Fanuc KAREL source: ka00105.KL

-- PROVISIONAL review KL for V940-1; original PC SHA256 45f8fe3be269b6ab01cad793c02046efcd257036997fb4219fc5ec4bbcc30542
-- Incomplete behavior may be omitted. Consult companion uncertainty JSON. Do not deploy.
PROGRAM KA00105
%NOLOCKGROUP
-- UNRESOLVED_DECL SRC type=000013
-- UNRESOLVED_DECL DST type=000013
BEGIN
  -- V9_ZERO_TABLE_METADATA_HINT layout=0001; no indexed target words; source/name/runtime held
  -- UNRESOLVED_PC offsets 5-20; opcodes 2E,22,32,35
  -- UNRESOLVED_PC offsets 25-40; opcodes 49,4A
  -- UNRESOLVED_PC offsets 45-49; opcodes 7F
END KA00105
